Fanuc KAREL source: kb00062.KL

-- PROVISIONAL review KL for V770-1; original PC SHA256 ebd9c32cf671465e3caa4a74d4ea210eae8f9b7b9a6a2028b338c7d584db132c
-- Incomplete behavior may be omitted. Consult companion uncertainty JSON. Do not deploy.
PROGRAM KB00062
%NOLOCKGROUP
BEGIN
  -- UNRESOLVED_PC offsets 5-12; opcodes 9D,23
  -- UNRESOLVED_PC offsets 17-27; opcodes 9D,22,9D,33,35
  -- UNRESOLVED_PC offsets 32-39; opcodes 9D,23
  -- UNRESOLVED_PC offsets 44-72; opcodes 27,22,22,22,22,31
  -- UNRESOLVED_PC offsets 77-81; opcodes 7F
END KB00062
